Fanuc KAREL source: kt00110.KL

-- PROVISIONAL review KL for V940-1; original PC SHA256 c8e20ec43066458ff6c2e9eea19d45ed5b0c94e0eac8862b9cfdda1a9514e07b
-- Incomplete behavior may be omitted. Consult companion uncertainty JSON. Do not deploy.
PROGRAM KT00110
%NOLOCKGROUP
VAR
  R1 : REAL
  OUT : REAL
-- UNRESOLVED_DECL Y2 type=002018
BEGIN
  -- V9_ZERO_TABLE_METADATA_HINT layout=0001; no indexed target words; source/name/runtime held
  -- UNRESOLVED_PC offsets 5-16; opcodes 2E,23
  -- UNRESOLVED_PC offsets 21-35; opcodes 2E,22,9D,33,B2
  -- UNRESOLVED_PC offsets 40-63; opcodes 21,22,9D,33,B1,64,6C,23
  -- UNRESOLVED_PC offsets 68-72; opcodes 7F
END KT00110
